// TIA Portal V20 export
Screen "MarriageFIFO_MB200_MB200RB04"  1260x525
  ScreenItem "Rectangle_4" at -3,2 size 1255x515  Type=HmiRectangle
  ScreenItem "Line_2" at 259,47 size 0x299  Type=HmiLine
  ScreenItem "Rectangle_6" at 4,5 size 1244x40  Type=HmiRectangle
  ScreenItem "Text_7" at 319,9 size 593x36  Type=HmiText
  ScreenItem "Faceplate container_1" at 3,47 size 1258x466  Type=HmiFaceplateContainer
